// TIA Portal V21 export
// export: Created 2026-10-12T11:32:14.3181651Z, ExportSetting WithDefaults, DisplayName Totally Integrated Automation Portal, DisplayVersion V21, DisplayName STEP 7 Professional, DisplayVersion V21, DisplayName STEP 7 Safety, DisplayVersion V21, DisplayName Tech WebApplication, DisplayVersion V21, DisplayName WinCC Basic/Comfort/Advanced, DisplayVersion V21, DisplayName WinCC Unified, DisplayVersion V21
FUNCTION "FC_OUTPUTS" : Void   // FC4, LAD
{ S7_Optimized_Access := 'TRUE' }
VERSION : 0.1
// stored: AutoNumber true, IsIECCheckEnabled false, SetENOAutomatically false, UDAEnableTagReadback false
BEGIN

REGION Network 1: CONVEYOR FWD ON
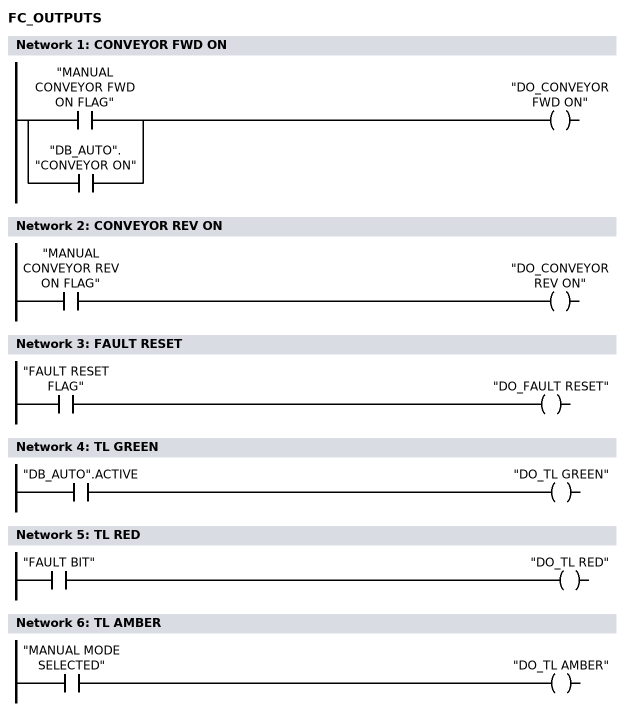
   RUNG wire#powerrail
      Contact( "MANUAL CONVEYOR FWD ON FLAG" )
      wire#w1
      Coil( "DO_CONVEYOR FWD ON" )
   END_RUNG
   RUNG wire#powerrail
      Contact( "DB_AUTO"."CONVEYOR ON" )
   END_RUNG wire#w1
   // the same network as SCL:
   "DO_CONVEYOR FWD ON" := "MANUAL CONVEYOR FWD ON FLAG" OR "DB_AUTO"."CONVEYOR ON";
END_REGION

REGION Network 2: CONVEYOR REV ON
   RUNG wire#powerrail
      Contact( "MANUAL CONVEYOR REV ON FLAG" )
      Coil( "DO_CONVEYOR REV ON" )
   END_RUNG
   // the same network as SCL:
   "DO_CONVEYOR REV ON" := "MANUAL CONVEYOR REV ON FLAG";
END_REGION

REGION Network 3: FAULT RESET
   RUNG wire#powerrail
      Contact( "FAULT RESET FLAG" )
      Coil( "DO_FAULT RESET" )
   END_RUNG
   // the same network as SCL:
   "DO_FAULT RESET" := "FAULT RESET FLAG";
END_REGION

REGION Network 4: TL GREEN
   RUNG wire#powerrail
      Contact( "DB_AUTO".ACTIVE )
      Coil( "DO_TL GREEN" )
   END_RUNG
   // the same network as SCL:
   "DO_TL GREEN" := "DB_AUTO".ACTIVE;
END_REGION

REGION Network 5: TL RED
   RUNG wire#powerrail
      Contact( "FAULT BIT" )
      Coil( "DO_TL RED" )
   END_RUNG
   // the same network as SCL:
   "DO_TL RED" := "FAULT BIT";
END_REGION

REGION Network 6: TL AMBER
   RUNG wire#powerrail
      Contact( "MANUAL MODE SELECTED" )
      Coil( "DO_TL AMBER" )
   END_RUNG
   // the same network as SCL:
   "DO_TL AMBER" := "MANUAL MODE SELECTED";
END_REGION
END_FUNCTION
